Fanuc KAREL source: kt00406.KL

-- PROVISIONAL review KL for V1013-1; original PC SHA256 b691edd8f408732d4bf6c29c1525b1584fe3ec6d26d871a26306cf675db03368
-- Incomplete behavior may be omitted. Consult companion uncertainty JSON. Do not deploy.
PROGRAM KT00406
%NOLOCKGROUP
VAR
  R1 : REAL
  R2 : REAL
  OUT : BOOLEAN
BEGIN
  -- UNRESOLVED_PC offsets 5-16; opcodes 2E,23
  -- UNRESOLVED_PC offsets 21-32; opcodes 2E,23
  -- UNRESOLVED_PC offsets 37-48; opcodes 2E,23
  -- UNRESOLVED_PC offsets 53-64; opcodes 2E,23
  -- UNRESOLVED_PC offsets 69-88; opcodes 21,21,71,23
  -- UNRESOLVED_PC offsets 93-97; opcodes 7F
END KT00406
